(* IEC 61131-3 sources: daoli-st-library/DL_Process (part 70) *)

(* ---- FB_DL_RecipeManager.st ---- *)
(*==============================================================================
 * 组件名称 (Component)  : FB_DL_RecipeManager
 * 所属子库 (Sublibrary) : DL_Process
 * 当前版本 (Version)    : 1.0.1
 * 兼容性 (Platform)   : CODESYS 3.5 / TwinCAT 3 / 汇川 InoProShop / Machine Expert
 *                         仅依赖 Standard.library（R_TRIG），零厂商方言
 * 分类     (Category)   : 工艺段功能块（Function Block · 通用配方管理器）
 * 功能简述 (Function)   : 以「参数清单 + 值集 + 校验和」承载多品种配方：选择、
 *                         校验、应用（写入运行参数）、写回（采集当前参数为
 *                         新配方）、切换防呆（仅机台稳态允许）、变更审计（次
 *                         数 + 注入时间戳）。零文件 I/O、零全局耦合——配方库
 *                         与运行参数均为引脚注入的数组，持久化由调用方自行完
 *                         成；校验和为自包含 32 位滚动异或累加，本块不伪造校
 *                         验和（写回时清零，由调用方重新生成）。
 * 首扫说明 (Init note)  : 纯事件型组件，免首扫（R23/公约 0.1），无 bInit；
 *                         所有状态由指令沿驱动。
 * 公约遵循 (Convention) : 0.2/R21 bError 为显式排除信息级码的派生式；0.4 双语
 *                         同行注释；0.5/R7 实例主体最前部无条件刷新；0.7/R15
 *                         故障锁存仅复位路径清码、信息级瞬时型；0.8 码位段
 *                         16#0005_xxxx（经 DL_Process VERSION.md 复核，本块
 *                         0140~0143 / 0240~0246 无冲突）；0.14 数组存取先判
 *                         域再索引、除法前判零（进度类运算无除法）；0.16 无
 *                         魔法数；0.17 终结符成对 ✓；0.18 ST_DL_RecipeEntry
 *                         与 E_DL_RecipeState 随本块同文件发布；0.19 码位同
 *                         行【级别】注释；0.20 验收向量入头注释；R25 bDone
 *                         单拍生命周期三律。
 * 红线自检 (Redline)    : R1 零全局变量表/外部变量引用 ✓｜R2 零物理 IO 地址 ✓
 *                         R3 纯 IEC 61131-3 ✓｜R4 越界/非有限值/校验和防御 ✓
 *                         R5 全变量中英双语同行注释 ✓｜R6 ENUM+CASE+ELSE ✓
 *                         R7 五实例（R_TRIG×4）主体最前部无条件刷新 ✓
 *                         R8 全常量化 ✓｜R25 单拍标志生命周期三律 ✓
 * 设计要点 (Key notes)  : ① 校验链（eValidating）：配方号域内 → 配方启用 →
 *                           参数个数一致 → 逐参数非有限值 → 逐参数上下限 →
 *                           校验和比对，任一失败锁存对应故障级码；
 *                         ② 应用（eApplying）单拍全量写入 afParamActual，防
 *                           半套参数生效；复核（eVerifying）回读重算校验和比
 *                           对，失败判写入异常 0245；
 *                         ③ 写回（Save）：运行参数拷入配方、个数同步、校验和
 *                           清零（本块不伪造校验和，调用方持久化前须重算）；
 *                         ④ 切换防呆：bMachineStopped=FALSE 时加载拒绝（信
 *                           息码 0141，不置故障，属正常联锁）；Load/Save 同
 *                           拍双丢弃（信息码 0142，"不猜"原则）；
 *                         ⑤ bParamOutOfRange 为瞬时型每拍重算（对当前选中配
 *                           方值集逐参数复核上下限），nOutOfRangeIndex 指向
 *                           首个越界参数；
 *                         ⑥ 数组维度字面量 16（等同 DL_RECIPE_MAX_PARAM）/32
 *                           （等同 DL_RECIPE_MAX_COUNT）与常量同步维护（跨
 *                           平台数组维度须编译期字面量，运行期域检查用常量）。
 * 偏离留档 (Deviation)  : 依 R11 头注释留档，共 1 条：
 *                         ① 校验和算法二选一裁定：规格允许复用 DL_Base 既有
 *                           CRC 函数或自包含算法；本块选自包含 32 位滚动异或
 *                           累加（uSum := (uSum XOR SHL(uSum,5)) +
 *                           REAL_TO_UDINT(v×1000.0 + 1.0E9)，正偏置保证折叠
 *                           项非负、避免负值参数取整的平台回绕歧义；取整语义
 *                           依平台四舍五入）。理由：保持本文件零跨子库依赖，
 *                           可单独导入；影响：与上层持久化校验格式必须一致
 *                           （调用方生成校验和时用同一含偏置算法），头注释已
 *                           声明。
 * 开源溯源 (Origin)     : 来源标签 codesys-forge / recipe-management
 *                         （RAW_NOTES_R8 S-6，T1-4 CODESYS Forge 首次开组：
 *                         公开配方管理示例——配方名/启用/参数值集/校验和的组
 *                         织分类与「校验→应用→复核」相语义，公开开源示例，
 *                         仅借鉴分类与参数域；结构体字段、状态机、码位、引脚
 *                         契约 100% 本库独立设计，clean-room 未复制源码。
 *                         许可证说明：借鉴对象为公开社区示例，本文件为本库原
 *                         创实现，随本库许可证发布）。
 * 验收向量 (Acceptance) :
 *   V1 正常 Load（3 参数，域内）→ bLoaded/eDone、uActiveChecksum 正确、
 *      uChangeCount +1、tLastChange 等于注入 tNow；
 *   V2 参数越界 → 故障 0243 + nOutOfRangeIndex 指向首个越界项；
 *   V3 校验和不匹配 → 0244（配方损坏）；
 *   V4 bMachineStopped=FALSE 加载 → 拒绝 + 信息码 0141（不置故障）；
 *   V5 Save 后 uChangeCount +1、配方值集与个数同步、uChecksum 清零；
 *   V6 Load+Save 同拍 → 双丢弃 + 信息码 0142；
 *   V7 配方参数含非有限值 → 0242；
 *   V8 配方号越界/未启用 → 0240。
 * 修订历史 (Revision)   :
 *   2026-11-15  v1.0.0  首版入库（Round 08 · DL_Process 配方管理件）
 *   2026-11-15  v1.0.1  R8 总监终审修复：终端态分支内的孤立空语句 `;`（非 IEC 61131-3 文法，statement_list 允许零条语句但不容纳孤立分号）改为纯注释占位分支，行为等价、跨平台可移植性合规。
 *============================================================================*)

(*-----------------------------------------------------------------------------
 * 结构体: ST_DL_RecipeEntry（归属 FB_DL_RecipeManager，与其同文件发布）
 *         值集维度字面量 16 等同 DL_RECIPE_MAX_PARAM，须与常量同步维护。
 *----------------------------------------------------------------------------*)
TYPE ST_DL_RecipeEntry :
STRUCT
    sName        : STRING[32];                    // 配方名（Recipe name）/ Recipe name
    bEnabled     : BOOL;                          // 配方启用（Enabled），FALSE 时选中即判故障 / Recipe enabled flag
    nParamCount  : UINT;                          // 有效参数个数（Active param count）[-]，域 0..16 / Active parameter count
    afValue      : ARRAY[0..15] OF REAL;          // 参数值集（Parameter values），维度 16 等同 DL_RECIPE_MAX_PARAM / Parameter values, dim 16
    uChecksum    : UDINT;                         // 校验和（Checksum），0=未启用校验；由调用方生成、本块只比对 / Checksum, 0 = verification off, caller generates
END_STRUCT
END_TYPE

(*-----------------------------------------------------------------------------
 * 枚举: E_DL_RecipeState（归属 FB_DL_RecipeManager，与其同文件发布）
 *----------------------------------------------------------------------------*)
TYPE E_DL_RecipeState :
(
    eIdle       := 0,   // 空闲：等操作沿 / Idle, awaiting operation edge
    eValidating := 10,  // 校验中：选择域/启用/个数/数值域/校验和逐项过链 / Validating selection, enable, count, ranges and checksum
    eApplying   := 20,  // 应用中：加载全量写入运行参数 / 写回采集参数入配方 / Applying, load writes parameters or save collects them
    eVerifying  := 30,  // 复核中：回读运行参数重算校验和比对 / Verifying, read-back checksum comparison
    eDone       := 40,  // 完成：结果保持，等下一操作沿 / Done, results held awaiting next operation
    eFault      := 99   // 故障锁存：仅复位沿退出 / Fault latched, only reset edge exits
) UINT;
END_TYPE

FUNCTION_BLOCK FB_DL_RecipeManager
VAR_INPUT
    bEnable             : BOOL;             // 使能（Enable），FALSE=中止操作并保持当前运行参数不变 / Enable, FALSE aborts and keeps live parameters
    bLoad               : BOOL;             // 加载所选配方到运行参数（Load），上升沿受理 / Load edge applies selected recipe
    bSave               : BOOL;             // 把当前运行参数写回所选配方（Save/Teach），上升沿受理 / Save edge teaches live parameters into recipe
    bValidate           : BOOL;             // 仅校验不应用（Validate），上升沿受理，结果出 bValid / Validate edge, result in bValid
    bMachineStopped     : BOOL := TRUE;     // 机台稳态确认（Machine stopped），FALSE 时拒绝加载（切换防呆）/ Machine stopped interlock, FALSE rejects load
    bReset              : BOOL;             // 复位故障（Fault reset），上升沿受理 / Rising edge resets fault
    nSelectRecipe       : UINT;             // 选中配方号（Selected recipe index）[-]，域 0..DL_RECIPE_MAX_COUNT-1 / Selected recipe index
    nParamCount         : UINT := 1;        // 本机参数个数（Param count）[-]，域 1..DL_RECIPE_MAX_PARAM，越界钳位 / Machine parameter count, clamped
    afParamMin          : ARRAY[0..15] OF REAL; // 参数下限（Param lower limits），逐项与配方值比较；min ≥ max 视为该参数未启用校验 / Param lower limits, min ≥ max disables that check
    afParamMax          : ARRAY[0..15] OF REAL; // 参数上限（Param upper limits），与下限配对使用 / Param upper limits paired with lower
    tNow                : TIME := T#0S;     // 时间戳注入（Timestamp injection）[ms]，禁读 CPU 钟，用于审计记录 / Injected timestamp for audit, CPU clock never read
END_VAR
VAR_OUTPUT
    bLoaded             : BOOL;             // 加载完成（Loaded），完成态且操作为 Load 时为 TRUE / TRUE while done with load operation
    bSaved              : BOOL;             // 写回完成（Saved），完成态且操作为 Save 时为 TRUE / TRUE while done with save operation
    bValid              : BOOL;             // 校验通过（Valid），校验型操作结果，保持到下次操作 / Validation verdict held until next operation
    bParamOutOfRange    : BOOL;             // 存在越界参数（Out of range），瞬时型每拍重算 / Transient out-of-range flag, recomputed each scan
    nOutOfRangeIndex    : UINT;             // 首个越界参数索引（First bad index）[-]，越界标志有效时成立 / First out-of-range parameter index
    nActiveRecipe       : UINT;             // 当前生效配方号（Active recipe）[-] / Currently applied recipe index
    uActiveChecksum     : UDINT;            // 当前运行参数校验和（Active checksum），每拍重算供上层比对 / Live parameter checksum recomputed each scan
    uChangeCount        : UDINT;            // 配方变更次数（Change counter），每次成功 Load/Save +1 / Successful load/save counter
    tLastChange         : TIME := T#0S;     // 末次变更时间戳（Last change time），取注入 tNow / Last change timestamp from injected tNow
    bBusy               : BOOL;             // 执行中（Busy），校验/应用/复核态为 TRUE / TRUE while validating/applying/verifying
    bDone               : BOOL;             // 操作完成单拍脉冲（Done pulse），单拍生命周期三律 / One-scan operation done pulse
    bError              : BOOL;             // 故障锁存（Error），仅故障级码置位 / Latched error, fault codes only
    uErrorId            : UDINT;            // 故障码（Error code），16#0005_xxxx 段，0=无故障 / Error code, fault-level priority
END_VAR
VAR_IN_OUT
    astRecipe           : ARRAY[0..31] OF ST_DL_RecipeEntry; // 配方库（Recipe library），维度 32 等同 DL_RECIPE_MAX_COUNT，调用方持有与持久化 / Recipe library owned and persisted by caller
    afParamActual       : ARRAY[0..15] OF REAL; // 当前运行参数（Live parameters），维度 16，Save 被读 / Load 被写 / Live parameters, read on save, written on load
END_VAR
VAR
    _eState             : E_DL_RecipeState := E_DL_RecipeState.eIdle; // 内部状态机（Internal state）/ Internal state
    _nOp                : USINT;            // 当前操作类型（Operation type）[-]，1=Load 2=Save 3=Validate，0=无 / Operation type register
    _bFaultLatch        : BOOL;             // 故障锁存标志（Fault latch flag），仅复位路径清除 / Fault latch, cleared only via reset path
    _uErrorIdInt        : UDINT;            // 内部故障级码寄存（Internal fault-level register）/ Internal fault-level register
    _uInfoCode          : UDINT;            // 本拍信息级码（Info code this cycle），瞬时型每拍重算 / Transient info code
    _nParamEff          : UINT;             // 生效参数个数（Effective param count），钳位后值 / Clamped effective parameter count
    _nSelEff            : UINT;             // 生效配方号（Effective recipe index），域校验后值 / Validated recipe index
    _fV                 : REAL;             // 循环内当前参数值（Loop value scratch）/ Loop parameter value scratch
    _bFinite            : BOOL;             // 非有限值检测结果（Finite check verdict）/ Finite-value check verdict
    _uSum               : UDINT;            // 校验和累加器（Checksum accumulator）/ Checksum accumulator
    _uTargetCk          : UDINT;            // 目标配方校验和（Target recipe checksum）/ Target recipe checksum
    _nIdx               : UINT;             // 循环索引（Loop index）[-] / Loop index
    _bBadIdxFound       : BOOL;             // 越界首索引已记录（First bad index found）/ First bad index recorded flag
    _bValOk             : BOOL;             // 校验链通过（Validation chain passed）/ Validation chain verdict
    _fbTrigLoad         : R_TRIG;           // 加载沿（Load edge detector）/ Load edge detector
    _fbTrigSave         : R_TRIG;           // 写回沿（Save edge detector）/ Save edge detector
    _fbTrigValidate     : R_TRIG;           // 校验沿（Validate edge detector）/ Validate edge detector
    _fbTrigReset        : R_TRIG;           // 复位沿（Reset edge detector）/ Reset edge detector
END_VAR
VAR CONSTANT
    DL_RECIPE_MAX_PARAM : UINT := 16;       // 单配方参数上限（Max params per recipe）[-]，与数组维度字面量 16 同步 / Max params, sync with literal dim 16
    DL_RECIPE_MAX_COUNT : UINT := 32;       // 配方库容量上限（Max recipe count）[-]，与数组维度字面量 32 同步 / Max recipes, sync with literal dim 32
    DL_RECIPE_REAL_MAX  : REAL := 3.4E38;   // 单精度有限值判据幅值（Finite magnitude bound），超出或非数均拒绝 / Finite magnitude bound for REAL inputs
    DL_RECIPE_EPS       : REAL := 1.0E-6;   // 浮点通用容差（General float epsilon）/ General float epsilon
    DL_RECIPE_VERIFY_EPS: REAL := 1.0E-3;   // 复核逐参数容差（Verify per-param epsilon），千分之一工程单位 / Verify tolerance per parameter
    DL_RECIPE_SCALE     : REAL := 1000.0;   // 校验和定标系数（Checksum scale）[-]，值×此系数取整入校验和 / Checksum scale factor for fixed-point fold
    DL_RECIPE_BIAS      : REAL := 1.0E9;    // 校验和正偏置（Checksum positive bias），保证折叠项非负、跨平台回绕确定 / Positive bias keeps fold term non-negative, portable
    DL_RECIPE_CHK_ROL   : DINT := 5;        // 校验和滚动移位量（Checksum shift amount）[-] / Checksum rolling shift amount
    DL_RECIPE_OP_LOAD   : USINT := 1;       // 操作码：加载（Op code: load）/ Op code load
    DL_RECIPE_OP_SAVE   : USINT := 2;       // 操作码：写回（Op code: save）/ Op code save
    DL_RECIPE_OP_VALID  : USINT := 3;       // 操作码：仅校验（Op code: validate only）/ Op code validate-only
    DL_RECIPE_ERR_SEL   : UDINT := 16#0005_0240; // 0005_0240 配方号越界/未启用【故障级】/ Bad recipe index or disabled, fault level
    DL_RECIPE_ERR_CNT   : UDINT := 16#0005_0241; // 0005_0241 参数个数与配方定义不一致【故障级】/ Param count mismatch, fault level
    DL_RECIPE_ERR_NAN   : UDINT := 16#0005_0242; // 0005_0242 配方参数含非有限值【故障级】/ Non-finite recipe parameter, fault level
    DL_RECIPE_ERR_RANGE : UDINT := 16#0005_0243; // 0005_0243 参数越界【故障级】/ Parameter out of range, fault level
    DL_RECIPE_ERR_CKSUM : UDINT := 16#0005_0244; // 0005_0244 校验和不匹配（配方损坏）【故障级】/ Checksum mismatch, recipe corrupted, fault level
    DL_RECIPE_ERR_VERIFY: UDINT := 16#0005_0245; // 0005_0245 应用后复核失败【故障级】/ Post-apply verify failed, fault level
    DL_RECIPE_ERR_STATE : UDINT := 16#0005_0246; // 0005_0246 非法状态兜底【故障级】/ Illegal state fallback, fault level
    DL_RECIPE_INFO_NOCK : UDINT := 16#0005_0140; // 0005_0140 配方未启用校验和（uChecksum=0）【信息级】/ Checksum disabled (zero), info level
    DL_RECIPE_INFO_LOCK : UDINT := 16#0005_0141; // 0005_0141 机台非稳态，加载被拒【信息级】/ Load rejected, machine not stopped, info level
    DL_RECIPE_INFO_CONF : UDINT := 16#0005_0142; // 0005_0142 Load/Save 同拍冲突，双丢弃【信息级】/ Load/save edge conflict, both dropped, info level
    DL_RECIPE_INFO_CLAMP: UDINT := 16#0005_0143; // 0005_0143 参数个数越界钳位【信息级】/ Param count clamped, info level
END_VAR

// ============================================================================
// 段 1｜实例无条件周期刷新（R7/0.5：严禁置于 IF/CASE 分支内）
//      Unconditional per-cycle refresh of all instances (R7/0.5)
// ============================================================================
_fbTrigLoad(CLK := bLoad);              // 加载沿（Load edge）
_fbTrigSave(CLK := bSave);              // 写回沿（Save edge）
_fbTrigValidate(CLK := bValidate);      // 校验沿（Validate edge）
_fbTrigReset(CLK := bReset);            // 复位沿（Reset edge）

// ============================================================================
// 段 2｜信息级预清零 + 单拍标志预清零 + 参数防御（R25/R15）
//      Info preset + one-shot preset + parameter defense (R25/R15)
// ============================================================================
_uInfoCode := 0;                        // 信息级瞬时型每拍重算（Transient info recomputed each scan）
bDone := FALSE;                         // 完成单拍先清零（R25：置位-消费-复位同周期闭环）/ Done pulse preset FALSE (R25 lifecycle)

// 参数个数钳位（Param count clamp，域 1..16）
IF nParamCount < UINT#1 THEN
    _nParamEff := UINT#1;               // 下限钳位（Lower clamp）
    _uInfoCode := DL_RECIPE_INFO_CLAMP; // 0005_0143 参数个数越界钳位【信息级】/ Count clamped, info level
ELSIF nParamCount > DL_RECIPE_MAX_PARAM THEN
    _nParamEff := DL_RECIPE_MAX_PARAM;  // 上限钳位（Upper clamp）
    _uInfoCode := DL_RECIPE_INFO_CLAMP; // 0005_0143 参数个数越界钳位【信息级】/ Count clamped, info level
ELSE
    _nParamEff := nParamCount;          // 引脚原值（Pin value as-is）
END_IF

// 复位路径：仅此路径可清故障锁存（R15）
IF _fbTrigReset.Q THEN
    _bFaultLatch := FALSE;              // 故障锁存解除（Fault latch released）
    _uErrorIdInt := 16#0000_0000;       // 故障码清零（Fault code cleared）
    IF _eState = E_DL_RecipeState.eFault THEN
        _eState := E_DL_RecipeState.eIdle; // 故障态回空闲（Fault state back to idle）
    END_IF
END_IF

// ============================================================================
// 段 3｜每拍瞬态复核：运行参数校验和 + 越界扫描（对当前选中配方）
//      Per-scan transient: live checksum + out-of-range scan on selected recipe
// ============================================================================
uActiveChecksum := 16#0000_0000;        // 校验和累加器清零（Checksum accumulator reset）
FOR _nIdx := UINT#0 TO _nParamEff - UINT#1 DO
    _fV := afParamActual[_nIdx];        // 索引域已由 _nParamEff 钳位保证（Index bounded by clamped count）
    uActiveChecksum := (uActiveChecksum XOR SHL(uActiveChecksum, DL_RECIPE_CHK_ROL))
                  + REAL_TO_UDINT(_fV * DL_RECIPE_SCALE + DL_RECIPE_BIAS);   // 滚动异或累加 + 正偏置保证非负折叠（偏离留档①算法）/ Rolling XOR fold with positive bias (deviation 1)
END_FOR

bParamOutOfRange := FALSE;              // 越界标志瞬态预清零（Transient flag preset）
nOutOfRangeIndex := UINT#0;             // 首个越界索引预清零（First bad index preset）
IF nSelectRecipe < DL_RECIPE_MAX_COUNT THEN
    IF (astRecipe[nSelectRecipe].nParamCount >= UINT#1)
      AND (astRecipe[nSelectRecipe].nParamCount <= DL_RECIPE_MAX_PARAM) THEN
        FOR _nIdx := UINT#0 TO astRecipe[nSelectRecipe].nParamCount - UINT#1 DO
            _fV := astRecipe[nSelectRecipe].afValue[_nIdx];      // 配方值（Recipe value）
            IF (afParamMin[_nIdx] < afParamMax[_nIdx])
              AND ((_fV < afParamMin[_nIdx]) OR (_fV > afParamMax[_nIdx]))
              AND (NOT bParamOutOfRange) THEN
                bParamOutOfRange := TRUE;            // 越界成立（Out of range found）
                nOutOfRangeIndex := _nIdx;           // 首个越界索引（First bad index）
            END_IF
        END_FOR
    END_IF
END_IF

// ============================================================================
// 段 4｜操作受理（仅在空闲/完成态受理指令沿；同拍冲突双丢弃）
//      Operation acceptance at idle/done; same-cycle conflict drops both
// ============================================================================
IF bEnable AND (( _eState = E_DL_RecipeState.eIdle)
             OR (_eState = E_DL_RecipeState.eDone)) THEN
    IF _fbTrigLoad.Q AND _fbTrigSave.Q THEN
        _uInfoCode := DL_RECIPE_INFO_CONF;  // 0005_0142 Load/Save 同拍冲突双丢弃【信息级】/ Edge conflict, both dropped
    ELSIF _fbTrigLoad.Q THEN
        IF bMachineStopped THEN
            _nOp := DL_RECIPE_OP_LOAD;      // 登记加载操作（Register load operation）
            _eState := E_DL_RecipeState.eValidating;
        ELSE
            _uInfoCode := DL_RECIPE_INFO_LOCK; // 0005_0141 机台非稳态加载被拒【信息级】/ Load rejected, machine running
        END_IF
    ELSIF _fbTrigSave.Q THEN
        _nOp := DL_RECIPE_OP_SAVE;          // 登记写回操作（Register save operation）
        _eState := E_DL_RecipeState.eValidating;
    ELSIF _fbTrigValidate.Q THEN
        _nOp := DL_RECIPE_OP_VALID;         // 登记校验操作（Register validate operation）
        _eState := E_DL_RecipeState.eValidating;
    END_IF
END_IF

// ============================================================================
// 段 5｜核心状态机（ENUM + CASE，含 ELSE 非法状态兜底）
//      Core state machine (ENUM + CASE with ELSE fallback)
// ============================================================================
CASE _eState OF

    E_DL_RecipeState.eIdle: // 空闲：等操作沿（受理逻辑在段 4）
        // 无动作（No action）

    E_DL_RecipeState.eValidating: // 校验链：域 → 启用 → 个数 → 非有限值 → 上下限 → 校验和
        _bValOk := TRUE;                    // 校验链初始通过（Chain starts valid）
        // ① 配方号域内（Index in domain）
        IF nSelectRecipe >= DL_RECIPE_MAX_COUNT THEN
            _bValOk := FALSE;
            _bFaultLatch := TRUE;
            _uErrorIdInt := DL_RECIPE_ERR_SEL;   // 0005_0240 配方号越界【故障级】/ Bad recipe index, fault level
        ELSE
            _nSelEff := nSelectRecipe;           // 生效配方号登记（Register effective index）
            // ② 配方启用（Recipe enabled）
            IF NOT astRecipe[_nSelEff].bEnabled THEN
                _bValOk := FALSE;
                _bFaultLatch := TRUE;
                _uErrorIdInt := DL_RECIPE_ERR_SEL; // 0005_0240 配方未启用【故障级】/ Recipe disabled, fault level
            END_IF
        END_IF

        IF _bValOk THEN
            // ③ 参数个数一致（Load/Validate 要求；Save 允许覆盖定义）
            IF (_nOp <> DL_RECIPE_OP_SAVE)
              AND (astRecipe[_nSelEff].nParamCount <> _nParamEff) THEN
                _bValOk := FALSE;
                _bFaultLatch := TRUE;
                _uErrorIdInt := DL_RECIPE_ERR_CNT;   // 0005_0241 个数与配方定义不一致【故障级】/ Count mismatch, fault level
            END_IF
        END_IF

        IF _bValOk AND (_nOp <> DL_RECIPE_OP_SAVE) THEN
            _uTargetCk := 16#0000_0000;          // 目标校验和累加器（Target checksum accumulator）
            FOR _nIdx := UINT#0 TO _nParamEff - UINT#1 DO
                _fV := astRecipe[_nSelEff].afValue[_nIdx];    // 配方值（Recipe value）
                _bFinite := (_fV >= (-DL_RECIPE_REAL_MAX)) AND (_fV <= DL_RECIPE_REAL_MAX); // 非有限值自比等价式（Finite check）
                IF NOT _bFinite THEN
                    _bValOk := FALSE;
                    _bFaultLatch := TRUE;
                    _uErrorIdInt := DL_RECIPE_ERR_NAN;        // 0005_0242 参数含非有限值【故障级】/ Non-finite parameter, fault level
                ELSIF (afParamMin[_nIdx] < afParamMax[_nIdx])
                  AND ((_fV < afParamMin[_nIdx]) OR (_fV > afParamMax[_nIdx])) THEN
                    _bValOk := FALSE;
                    _bFaultLatch := TRUE;
                    _uErrorIdInt := DL_RECIPE_ERR_RANGE;      // 0005_0243 参数越界【故障级】/ Parameter out of range, fault level
                    nOutOfRangeIndex := _nIdx;                // 首个越界索引（First bad index）
                END_IF
                _uTargetCk := (_uTargetCk XOR SHL(_uTargetCk, DL_RECIPE_CHK_ROL))
                         + REAL_TO_UDINT(_fV * DL_RECIPE_SCALE + DL_RECIPE_BIAS);   // 同算法重算目标校验和（Target checksum recomputed, same algorithm）
            END_FOR
            // ⑤ 校验和比对（=0 视为未启用校验）
            IF _bValOk THEN
                IF astRecipe[_nSelEff].uChecksum = 16#0000_0000 THEN
                    _uInfoCode := DL_RECIPE_INFO_NOCK;    // 0005_0140 未启用校验和【信息级】/ Checksum disabled, info level
                ELSIF astRecipe[_nSelEff].uChecksum <> _uTargetCk THEN
                    _bValOk := FALSE;
                    _bFaultLatch := TRUE;
                    _uErrorIdInt := DL_RECIPE_ERR_CKSUM;  // 0005_0244 校验和不匹配（配方损坏）【故障级】/ Checksum mismatch, fault level
                END_IF
            END_IF
        END_IF

        // 校验链出口分派（Chain exit dispatch）
        IF _bValOk THEN
            IF _nOp = DL_RECIPE_OP_LOAD THEN
                _eState := E_DL_RecipeState.eApplying;    // 进入应用（Proceed to apply）
            ELSIF _nOp = DL_RECIPE_OP_SAVE THEN
                _eState := E_DL_RecipeState.eApplying;    // 写回也走应用相（Save proceeds to apply phase）
            ELSE
                bValid := TRUE;                           // 仅校验：结果通过（Validate-only passed）
                bDone := TRUE;                            // 完成单拍（R25 本拍闭环）/ Done pulse (R25)
                _eState := E_DL_RecipeState.eDone;
            END_IF
        ELSE
            _eState := E_DL_RecipeState.eFault;           // 校验失败进故障锁存（Validation failed, latch fault）
        END_IF

    E_DL_RecipeState.eApplying: // 应用：Load 单拍全量写入 / Save 单拍全量采集
        IF _nOp = DL_RECIPE_OP_LOAD THEN
            FOR _nIdx := UINT#0 TO _nParamEff - UINT#1 DO
                _fV := astRecipe[_nSelEff].afValue[_nIdx];    // 源：配方值（Source: recipe value）
                _bFinite := (_fV >= (-DL_RECIPE_REAL_MAX)) AND (_fV <= DL_RECIPE_REAL_MAX);
                IF _bFinite THEN
                    afParamActual[_nIdx] := _fV;              // 单拍全量写入（Single-scan bulk write, no half-set applied）
                END_IF
            END_FOR
            _eState := E_DL_RecipeState.eVerifying;           // 进入复核（Proceed to verify）
        ELSE
            FOR _nIdx := UINT#0 TO _nParamEff - UINT#1 DO
                astRecipe[_nSelEff].afValue[_nIdx] := afParamActual[_nIdx]; // 单拍全量采集（Single-scan bulk collect）
            END_FOR
            astRecipe[_nSelEff].nParamCount := _nParamEff;    // 个数同步（Count synchronized）
            astRecipe[_nSelEff].uChecksum := 16#0000_0000;    // 校验和清零：本块不伪造，调用方须重算（Checksum zeroed, caller regenerates）
            uChangeCount := uChangeCount + UINT#1;            // 审计计数（Audit counter）
            tLastChange := tNow;                              // 审计时间戳取注入值（Audit timestamp from injected pin）
            nActiveRecipe := _nSelEff;                        // 生效配方号登记（Active recipe registered）
            bSaved := TRUE;                                   // 写回完成保持（Saved held）
            bDone := TRUE;                                    // 完成单拍（R25 本拍闭环）/ Done pulse (R25)
            _eState := E_DL_RecipeState.eDone;
        END_IF

    E_DL_RecipeState.eVerifying: // 复核：回读运行参数与目标比对（防写入异常）
        IF astRecipe[_nSelEff].uChecksum <> 16#0000_0000 THEN
            IF uActiveChecksum <> astRecipe[_nSelEff].uChecksum THEN
                _bFaultLatch := TRUE;
                _uErrorIdInt := DL_RECIPE_ERR_VERIFY;         // 0005_0245 复核失败（写入异常）【故障级】/ Verify failed, fault level
                _eState := E_DL_RecipeState.eFault;
            ELSE
                nActiveRecipe := _nSelEff;                    // 生效配方号登记（Active recipe registered）
                uChangeCount := uChangeCount + UINT#1;        // 审计计数（Audit counter）
                tLastChange := tNow;                          // 审计时间戳（Audit timestamp）
                bLoaded := TRUE;                              // 加载完成保持（Loaded held）
                bDone := TRUE;                                // 完成单拍（R25 本拍闭环）/ Done pulse (R25)
                _eState := E_DL_RecipeState.eDone;
            END_IF
        ELSE
            // 目标未启用校验和：逐参数容差比对兜底（Checksum off: element-wise tolerance fallback）
            FOR _nIdx := UINT#0 TO _nParamEff - UINT#1 DO
                IF ABS(afParamActual[_nIdx] - astRecipe[_nSelEff].afValue[_nIdx]) > DL_RECIPE_VERIFY_EPS THEN
                    _bFaultLatch := TRUE;
                    _uErrorIdInt := DL_RECIPE_ERR_VERIFY;     // 0005_0245 复核失败【故障级】/ Verify failed, fault level
                    _eState := E_DL_RecipeState.eFault;
                END_IF
            END_FOR
            IF NOT _bFaultLatch THEN
                nActiveRecipe := _nSelEff;
                uChangeCount := uChangeCount + UINT#1;
                tLastChange := tNow;
                bLoaded := TRUE;                              // 加载完成保持（Loaded held）
                bDone := TRUE;                                // 完成单拍（R25）/ Done pulse (R25)
                _eState := E_DL_RecipeState.eDone;
            END_IF
        END_IF

    E_DL_RecipeState.eDone: // 完成：结果保持，下一操作沿回空闲（受理逻辑在段 4，下一拍起效）
        IF _fbTrigLoad.Q OR _fbTrigSave.Q OR _fbTrigValidate.Q THEN
            _eState := E_DL_RecipeState.eIdle;                // 让位新操作（Yield to new operation）
            bLoaded := FALSE;                                 // 结果锁存随让位清零（Result holds released）
            bSaved := FALSE;
            bValid := FALSE;
        END_IF

    E_DL_RecipeState.eFault: // 故障锁存：等复位（复位路径在段 2）
        // 等复位（Awaiting reset）

    ELSE // 非法状态兜底（本块专用码位）
        _bFaultLatch := TRUE;
        _uErrorIdInt := DL_RECIPE_ERR_STATE;                  // 0005_0246 非法状态兜底【故障级】/ Illegal state fallback, fault level
        _eState := E_DL_RecipeState.eFault;
END_CASE

// ============================================================================
// 段 6｜使能撤销与出口派生（R21）
//      Enable teardown and outlet derivation (R21)
// ============================================================================
IF NOT bEnable THEN
    // 撤销进行中操作，运行参数保持不变（Abort in-flight ops, live parameters untouched）
    IF (_eState = E_DL_RecipeState.eValidating)
     OR (_eState = E_DL_RecipeState.eApplying)
     OR (_eState = E_DL_RecipeState.eVerifying) THEN
        _eState := E_DL_RecipeState.eIdle;   // 中途回空闲（Back to idle mid-flight）
    END_IF
END_IF

bBusy := (_eState = E_DL_RecipeState.eValidating)
      OR (_eState = E_DL_RecipeState.eApplying)
      OR (_eState = E_DL_RecipeState.eVerifying);            // 执行中派生（Busy derived）

bError := _bFaultLatch;                      // 故障级派生式（Fault-level derived form）
IF _bFaultLatch THEN
    uErrorId := _uErrorIdInt;                // 故障级码优先透出（Fault-level priority）
ELSE
    uErrorId := _uInfoCode;                  // 无故障时透出本拍信息级码（Transient info code）
END_IF
END_FUNCTION_BLOCK

(* ---- FB_DL_RejectBlowCtrl.st ---- *)
(*
    FB_DL_RejectBlowCtrl —— 输送线剔除气吹执行时序（NG 预告 → 距离/速度延时 → 定宽气吹 → 对账）
    ------------------------------------------------------------------
    组件名称  : FB_DL_RejectBlowCtrl
    分类      : DL_Process / Rejection
    前缀      : FB_DL_
    版本      : 1.0.0
    溯源      : 自研线 s9-conv（R7 先例同口径）：剔除气吹执行时序属输送线
                工程惯例的 clean-room 自有实现；判定域（视觉 / 称重）与
                诊断域（堵塞）归邻件，本件零借用；实现 / 引脚名 / 码位 /
                对账口径 100% 自有；无闭源参考。
    平台      : 纯 IEC 61131-3（ENUM + CASE + TON / R_TRIG + 标准换算），
                CODESYS 3.5 / TwinCAT 3 / InoProShop / Machine Expert 通用
    作者      : 道莅代码库 · PLC编程专家（R72 构建轮 · 批 4 · 序号 11）
    ------------------------------------------------------------------
    功能说明  : 灌装 / 包装线吹除 NG 瓶：eIdle →（bNgFlag 上升沿布防）
                eArm（延时窗 = fDistNgToGate / fBeltVel 秒换算毫秒，组态
                容差即引脚侧自行加权，本件按纯行程 / 速度口径）→ eBlow
                （定宽气吹脉冲 tBlowPulse）→ eConfirm（确认窗 tConfirmWin
                满拍**复验一次** NG 离线状态，R41/R42 同拍竞态口径：窗满拍
                反馈迟到临界收敛以窗满拍采样为准）→ eIdle。
                对账口径（漏剔 / 误剔 / 剔除三值互斥，窗满拍一次性判归）：
                ① 漏剔 uMissCount：窗满拍 bNgFlag 仍在位（气吹未吹走 NG）；
                ② 误剔 uFalseCount：布防后气吹执行拍 bNgFlag 已离线（无 NG
                   确认却执行气吹——预告为伪沿，好品被吹）；
                ③ 剔除 uRejectCount：气吹拍 NG 在位且窗满拍已离线（正常剔除）。
                漏剔 / 误剔计数直接进 OEE 质量因子。
                安全口径：
                ① fBeltVel 非有限 / <= 0 → **拒收布防 + NG 漏剔计数**（不发
                   气吹，防静默放行——速度不明即不剔除，宁可人工清台），
                   信息级；执行中途速度失效同样撤销布防 + 漏剔计数；
                ② 除法先判后除：fDistNgToGate / fBeltVel 仅在速度过闸后执行；
                   毫秒换算 LREAL→DINT 前做实数上界钳制（DL_RBC_TMAX，
                   防溢出方向翻转，R151）；
                ③ 失能 → bBlowCmd 清零 + 布防撤销（停机相输出清零，R57）；
                   计数保留（OEE 台账语义）；
                ④ 组态闸：tBlowPulse / tConfirmWin 非正 或 fDistNgToGate
                   非有限 / 非正 → 故障锁存（锁存期 NG 沿一律按漏剔计数，
                   宁多计不漏计）。
    错误码    : 16#0005_0630 速度不明拒剔（fBeltVel 非有限 / 非正，布防撤销
                            + 漏剔计数），条件期重算 —— 信息级，不置 bError
                16#0005_0631 组态非法（tBlowPulse / tConfirmWin 非正 /
                            fDistNgToGate 非有限 / 非正），锁存至复位沿
                            —— 故障级
                加码反证句（R90）：0630 由「布防撤销 + 漏剔计数递增」唯一
                观测（正常剔除路径漏剔计数不动）；0631 与 0630 输出可分
                （bError 与锁存回放 vs 条件信息级），成因互斥（组态表 vs
                运行速度），故各立一码。
    码位总账  : 16#0005_0630 用 ｜ 16#0005_0631 用
                （0620~0622 / 3036~3038 已由同段邻件占用，本件不占）
    边界与披露: 一 R_TRIG（rtNg / rtReset）与 TON（tonPhase）每拍**无条件
                   调用**（规则 ⑦）；tonPhase PT 按相选择（布防延时 / 气吹
                   定宽 / 确认窗三态一实例，R367 逐相 PT 口径），IN = 相驻留
                   显式变量；
                二 零全局变量、零 VAR_EXTERNAL、零物理地址；
                三 归属 Ownership：E_DL_RejectPhase 属主为本文件（全库唯一
                   定义，R264），引用件只引用不重声明；
                四 状态机 ENUM + CASE 必带 ELSE 兜底（非法枚举值 → eFault
                   锁存）+ 段 5b 统一故障迁入闸（R274）；
                五 域闸逐项点名（R272）：fBeltVel / fDistNgToGate 双浮点引脚
                   全部纳入非有限与符号闸；
                六 换算链：tArmDelay := DINT_TO_TIME(LREAL_TO_DINT(钳制后的
                   行程毫秒))，钳制上界 2147483000 ms（< 2^31 − 347，
                   LREAL_TO_DINT 域内可表反算，R63）；
                七 分工声明：FB_DL_VisionResultGate（视觉结果放行闸）、
                   FB_DL_WeightCheckReject（称重 NG 判定）、
                   FB_DL_ConveyorJamDetect（堵塞诊断）——三者均属「判定」域，
                   本件只做「预告 → 延时 → 气吹 → 对账」**执行时序**域
                   （R363 邻接共存先例），不判 NG、不诊断堵塞；
                八 复位沿作用域（R311）：清故障锁存 + 清锁存码 + 迁 eIdle +
                   撤布防，**不清** uRejectCount / uMissCount / uFalseCount
                   （OEE 台账语义，只随失能保留、由上位归档后清）；
                九 依赖声明：仅 Standard.library（TON / R_TRIG），零厂商
                   方言；
                十 接口契约：bNgFlag 须为**电平型**预告（预告对象离线前保持
                   在位），脉型预告会在气吹拍被判为误剔（uFalseCount 虚高）
                   ——脉型上游须先展宽再接入；失能相（bEn = FALSE）的 NG 沿
                   不布防不计数（停线工况，宁缺勿滥口径）。
    验收向量  : V1 正常剔除：NG 沿 → 行程延时 → 气吹拍 NG 在位 → 窗满拍
                NG 离线 → uRejectCount + 1；
                V2 漏剔：窗满拍 bNgFlag 仍在位 → uMissCount + 1；
                V3 误剔：气吹拍 bNgFlag 已离线 → uFalseCount + 1；
                V4 fBeltVel = 0 / NaN → NG 沿按漏剔计数、不发气吹、0630；
                V5 tBlowPulse = T#0MS → 0631 锁存；V6 失能 → bBlowCmd 清零
                + 布防撤销；V7 复位沿 → 解锁回 eIdle（计数不清）。
                算法已证（脚本）：未跑 ｜ 编译器已证（三平台）：未跑
    修订记录  : 2026-11-23 v1.0.0 首次入库（R72 构建轮 · 批 4 · 序号 11）
*)
TYPE E_DL_RejectPhase :
(
    eIdle    := 0,                         // 空闲：等 NG 预告沿布防 / idle, waiting for the NG leading edge
    eArm     := 10,                        // 布防延时：行程 / 速度换算延时窗 / armed, the travel delay window
    eBlow    := 20,                        // 定宽气吹：tBlowPulse 定宽脉冲 / blowing, the fixed width pulse
    eConfirm := 30,                        // 确认窗：窗满拍复验 NG 离线 / confirm, the recheck window
    eFault   := 60                         // 故障：锁存待复位 / fault, latched until the reset
);
END_TYPE

FUNCTION_BLOCK FB_DL_RejectBlowCtrl
VAR_INPUT
    bNgFlag       : BOOL := FALSE;         (* 上游 NG 预告（视觉 / 称重判定输出），[标志] / the upstream NG leading flag *)
    fBeltVel      : LREAL := 1000.0;       (* 输送带速度，[mm/s]，非有限或非正拒剔 / the belt velocity in mm per second *)
    fDistNgToGate : LREAL := 500.0;        (* NG 检测位到气吹位间距，[mm]，禁非有限 / 非正 / the distance from the detector to the gate in mm *)
    tBlowPulse    : TIME := T#100MS;       (* 气吹定宽，[ms]，禁非正 / the blow pulse width *)
    tConfirmWin   : TIME := T#200MS;       (* 剔除确认窗，[ms]，禁非正 / the reject confirmation window *)
    bEn           : BOOL := FALSE;         (* 使能，[标志]，FALSE 撤布防清气吹（计数保留）/ the enable *)
    bReset        : BOOL := FALSE;         (* 故障复位，[标志]，上升沿唯一解除 / the fault reset *)
END_VAR
VAR_OUTPUT
    bBlowCmd    : BOOL := FALSE;           (* 气吹指令出口（定宽脉冲），[标志] / the blow command outlet *)
    uRejectCount: UDINT := 0;              (* 剔除成功计数（OEE 台账），[件] / the successful reject count *)
    uMissCount  : UDINT := 0;              (* 漏剔计数（窗满 NG 仍在位 / 速度不明拒剔），[件] / the miss count *)
    uFalseCount : UDINT := 0;              (* 误剔计数（气吹拍 NG 已离线），[件] / the false reject count *)
    eState      : E_DL_RejectPhase := E_DL_RejectPhase.eIdle; // 主状态机当前态 [状态] / the current state
    bError      : BOOL := FALSE;           (* 故障标志，与锁存同源（R191）/ the fault flag from the latch *)
    nErrCode    : UDINT := 16#0000_0000;   (* 错误码，0 = 正常，故障锁存回放（R187）/ the error id *)
END_VAR
VAR
    _bInit      : BOOL := FALSE;           (* 首拍初始化标志（R310）/ the first scan flag *)
    _eState     : E_DL_RejectPhase := E_DL_RejectPhase.eIdle; // 内部状态寄存器 / the internal state register
    _bFault     : BOOL := FALSE;           (* 故障锁存副本，仅复位沿解除 / the fault latch copy *)
    _nCodeLatch : UDINT := 0;              (* 锁存成因码，故障期回放 / the latched cause code *)
    _bVelBad    : BOOL := FALSE;           (* 速度不明标志（逐拍重算，R272 闸）/ the velocity invalid flag *)
    _bCfgBad    : BOOL := FALSE;           (* 组态非法标志（逐拍重算，仅用于首次锁存）/ the config fault flag *)
    _bBlow      : BOOL := FALSE;           (* 气吹单相内部位（统一出口映射）/ the internal blow bit *)
    _bFalseSus  : BOOL := FALSE;           (* 误剔嫌疑标志（气吹拍 NG 已离线登记）/ the false reject suspect flag *)
    _tArmDelay  : TIME := T#0S;             (* 布防延时换算值（过闸后逐拍重算）[ms] / the computed arm delay *)
    _tPhasePt   : TIME := T#0S;             (* 逐相 PT 预置（R367：每拍先给缺省再按相覆盖）[ms] / the per phase PT preset *)
    _fDelayMs   : LREAL := 0.0;             (* 行程毫秒中间量（钳制前）[ms] / the travel milliseconds temporary *)
    nDelayMs    : DINT := 0;                (* 钳制后的行程毫秒 [ms] / the clamped travel milliseconds *)
    rtNg        : R_TRIG;                  (* NG 预告上升沿实例（无条件调用）/ the NG leading edge instance *)
    rtReset     : R_TRIG;                  (* 复位沿实例（无条件调用）/ the reset edge instance *)
    tonPhase    : TON;                     (* 相计时实例（逐相 PT，无条件调用，R367）/ the phase timer *)
    _bPhaseIn   : BOOL := FALSE;           (* 相驻留判据（tonPhase IN 显式变量）/ the phase residency flag *)
END_VAR
VAR CONSTANT
    DL_RBC_CODE_VEL : UDINT := 16#0005_0630; // 速度不明信息码 [码] / the velocity info code
    DL_RBC_CODE_CFG : UDINT := 16#0005_0631; // 组态非法故障码 [码] / the config fault code
    DL_RBC_TZERO    : TIME := T#0S;          (* 零时长哨兵 [ms] / the zero duration sentinel *)
    DL_RBC_TMAX     : LREAL := 2147483000.0; (* 换算毫秒钳制上界（< 2^31 可表反算，R63）[ms] / the conversion clamp ceiling *)
    DL_RBC_CMAX     : UDINT := 2147483000;   (* 计数饱和上限（UDINT 域，防回绕）[件] / the count saturation cap *)
    DL_RBC_MS_SEC   : LREAL := 1000.0;       (* 秒到毫秒换算常量乘子 [ms/s] / the seconds to milliseconds multiplier *)
    DL_RBC_FZERO    : LREAL := 0.0;          (* 浮点零哨兵 [mm/s 或 mm] / the float zero sentinel *)
    DL_RBC_ZERO     : UDINT := 0;            (* 无符号零哨兵 [码或件] / the unsigned zero sentinel *)
    DL_RBC_ONE      : UDINT := 1;            (* 计数步进 [件] / the count step *)
END_VAR

// 段 0｜沿检测无条件周期调用（规则 ⑦）/ segment 0, the unconditional edge refresh
rtNg(CLK := bNgFlag);                      // NG 预告沿 / the NG leading edge
rtReset(CLK := bReset);                    // 复位沿 / the reset edge

// 段 1｜首拍初始化（R310）/ segment 1, the first scan init
IF NOT _bInit THEN                         // 首拍一拍 / the first scan
    _bInit := TRUE;                        // 置首拍标志 / raise the first scan flag
    _bFault := FALSE;                      // 故障锁存显式清零 / clear the fault latch explicitly
    _eState := E_DL_RejectPhase.eIdle;     // 状态显式落空闲 / place the state to idle
END_IF

// 段 2｜域闸（R272 全枚举：fBeltVel / fDistNgToGate 双引脚；非有限双判 R79）/ segment 2, the domain gates
_bVelBad := (fBeltVel <> fBeltVel) OR ((fBeltVel - fBeltVel) <> DL_RBC_FZERO) OR (fBeltVel <= DL_RBC_FZERO); // 速度非有限或非正 / the velocity invalid
_bCfgBad := (tBlowPulse <= DL_RBC_TZERO) OR (tConfirmWin <= DL_RBC_TZERO) // 定宽或确认窗非正 / a non positive pulse or window
         OR (fDistNgToGate <> fDistNgToGate) OR ((fDistNgToGate - fDistNgToGate) <> DL_RBC_FZERO) // 间距非有限 / the distance non finite
         OR (fDistNgToGate <= DL_RBC_FZERO); // 间距非正 / a non positive distance

// 段 3｜复位沿与首次成因锁存（复位沿唯一解除，R188；故障期不重推断，R189）/ segment 3, the reset edge and the first cause latch
IF rtReset.Q THEN                          // 复位上升沿 / the reset rising edge
    _bFault := FALSE;                      // 清故障锁存（恒可达，R152 自证）/ clear the fault latch
    _nCodeLatch := DL_RBC_ZERO;            // 清锁存码（作用域 R311：不清三计数，台账语义）/ clear the latched code
    _eState := E_DL_RejectPhase.eIdle;     // 迁回空闲 / back to idle
END_IF
IF (NOT _bFault) AND _bCfgBad THEN         // 组态非法未锁存命中 / a config fault hit
    _bFault := TRUE;                       // 置锁存 / latch the fault
    _nCodeLatch := DL_RBC_CODE_CFG;        // 登记组态码 / register the config code
END_IF

// 段 4｜布防延时换算（先判后除：速度过闸才做除法；实数上界钳制防换算溢出）/ segment 4, the arm delay conversion
IF (NOT _bVelBad) AND (NOT _bCfgBad) THEN  // 双闸通过才换算 / both gates passed
    _fDelayMs := (fDistNgToGate / fBeltVel) * DL_RBC_MS_SEC; // 行程 / 速度 × 1000（除子已闸非零非有限）/ the travel milliseconds
    IF _fDelayMs > DL_RBC_TMAX THEN        // 实数上界钳制（防 LREAL_TO_DINT 溢出方向翻转，R151）/ the clamp before narrowing
        nDelayMs := LREAL_TO_DINT(DL_RBC_TMAX); // 钳到上界 / clamp to the ceiling
    ELSIF _fDelayMs < DL_RBC_FZERO THEN    // 负值防御（双闸后结构性不可达，兜底口径）/ the negative guard
        nDelayMs := 0;                     // 钳到零 / clamp to zero
    ELSE                                   // 域内换算 / the in domain conversion
        nDelayMs := LREAL_TO_DINT(_fDelayMs); // 标准降位转换 / the standard narrowing
    END_IF
    _tArmDelay := DINT_TO_TIME(nDelayMs);  // 毫秒转 TIME / the milliseconds to TIME
ELSE                                       // 闸未通过 / the gates failed
    _tArmDelay := DL_RBC_TZERO;            // 延时清零（布防路径已拒收）/ zero the delay
END_IF

// 段 5｜主状态机（ENUM + CASE，ELSE 兜底；相驻留显式变量供段 0b 定时器）/ segment 5, the main state machine
CASE _eState OF

    E_DL_RejectPhase.eIdle:                // 空闲相：等 NG 沿布防 / the idle phase
        _bBlow := FALSE;                   // 气吹位清零 / clear the blow bit
        IF rtNg.Q AND bEn AND (NOT _bFault) AND (NOT _bVelBad) AND (NOT _bCfgBad) THEN // 布防沿 + 全量闸位复检（R274）/ the arming edge with the full gate recheck
            _bFalseSus := FALSE;           // 布防清嫌疑标志 / clear the suspect flag
            _eState := E_DL_RejectPhase.eArm; // 迁入布防相 / enter the arm phase
        ELSIF rtNg.Q AND bEn AND (NOT _bFault) AND (_bVelBad OR _bCfgBad) THEN // 速度不明的 NG 沿（组态非法沿已在段 3 先锁存，不会进入本支）/ the NG edge with an invalid velocity
            IF uMissCount < DL_RBC_CMAX THEN // 饱和闸（UDINT 域防回绕）/ the saturation cap
                uMissCount := uMissCount + DL_RBC_ONE; // 漏剔计数（速度不明即不剔除，宁可人工清台）/ count a miss
            END_IF
        END_IF                             // 失能相的 NG 沿不布防不计数（停线工况声明，头注释边界十）

    E_DL_RejectPhase.eArm:                 // 布防相：等行程延时 / the arm phase
        IF (NOT bEn) OR _bVelBad THEN      // 失能或速度中途失效：撤布防 + 漏剔计数 / the disarm on disable or velocity loss
            IF uMissCount < DL_RBC_CMAX THEN // 饱和闸 / the saturation cap
                uMissCount := uMissCount + DL_RBC_ONE; // 漏剔计数 / count a miss
            END_IF
            _eState := E_DL_RejectPhase.eIdle; // 撤布防回空闲 / disarm to idle
        ELSIF tonPhase.Q THEN              // 行程延时计满（零延时换算合法，立即吹口径）/ the delay elapsed
            _eState := E_DL_RejectPhase.eBlow; // 迁入气吹相 / enter the blow phase
        END_IF

    E_DL_RejectPhase.eBlow:                // 气吹相：定宽脉冲 + 误剔登记 / the blow phase
        _bBlow := TRUE;                    // 气吹位置位 / raise the blow bit
        IF (NOT bNgFlag) AND (NOT _bFalseSus) THEN // NG 已离线却执行气吹（电平型预告伪沿，接口契约见头注释边界十）登记嫌疑（一次性）/ the false reject registration
            _bFalseSus := TRUE;            // 置嫌疑标志（窗满拍判归互斥用）/ raise the suspect flag
            IF uFalseCount < DL_RBC_CMAX THEN // 饱和闸 / the saturation cap
                uFalseCount := uFalseCount + DL_RBC_ONE; // 误剔计数（布防后无 NG 确认却执行气吹）/ count a false reject
            END_IF
        END_IF
        IF (NOT bEn) OR _bVelBad THEN      // 气吹中失能 / 速度失效：撤气吹（安全侧停吹）/ the blow abort
            _bBlow := FALSE;               // 气吹位清零 / clear the blow bit
            _eState := E_DL_RejectPhase.eIdle; // 回空闲 / to idle
        ELSIF tonPhase.Q THEN              // 定宽计满 / the pulse elapsed
            _bBlow := FALSE;               // 定宽到撤气吹（R129 两拍口径：本拍撤、映射段不再改）/ drop the blow bit
            _eState := E_DL_RejectPhase.eConfirm; // 迁入确认相 / enter the confirm phase
        END_IF

    E_DL_RejectPhase.eConfirm:             // 确认相：窗满拍复验一次（R41/R42：窗满拍采样为准）/ the confirm phase
        IF (NOT bEn) THEN                  // 失能：撤销对账（失能拍不判归，声明口径）/ the disabled confirm
            _eState := E_DL_RejectPhase.eIdle; // 回空闲 / to idle
        ELSIF tonPhase.Q THEN              // 确认窗满拍 / the window full scan
            IF bNgFlag THEN                // 窗满拍 NG 仍在位（气吹未吹走 NG）/ the NG still present
                IF uMissCount < DL_RBC_CMAX THEN // 饱和闸 / the saturation cap
                    uMissCount := uMissCount + DL_RBC_ONE; // 漏剔计数 / count a miss
                END_IF
            ELSIF NOT _bFalseSus THEN      // 窗满离线且非误剔嫌疑（气吹拍在位）→ 正常剔除判归 / the normal reject verdict
                IF uRejectCount < DL_RBC_CMAX THEN // 饱和闸 / the saturation cap
                    uRejectCount := uRejectCount + DL_RBC_ONE; // 剔除成功计数 / count a reject
                END_IF
            END_IF                         // 误剔嫌疑者已在气吹拍计入 uFalseCount，三值互斥不重复判归
            _bFalseSus := FALSE;           // 判归完成清嫌疑 / clear the suspect flag
            _eState := E_DL_RejectPhase.eIdle; // 回空闲 / to idle
        END_IF

    E_DL_RejectPhase.eFault:               // 故障相：等复位沿（解除可达）；锁存期 NG 沿按漏剔计数（宁多计不漏计，码位声明口径）/ the fault phase with the miss accounting
        IF rtNg.Q AND bEn THEN             // 锁存期 NG 沿 / the NG edge while latched
            IF uMissCount < DL_RBC_CMAX THEN // 饱和闸 / the saturation cap
                uMissCount := uMissCount + DL_RBC_ONE; // 漏剔计数 / count a miss
            END_IF
        END_IF
        IF NOT _bFault THEN                // 锁存已清才迁出 / the exit after the latch cleared
            _eState := E_DL_RejectPhase.eIdle; // 迁回空闲 / back to idle
        END_IF

    ELSE                                   // 非法枚举值拦截 / the illegal enumeration guard
        _eState := E_DL_RejectPhase.eFault; // 落故障相 / force to the fault phase
        _bFault := TRUE;                   // 置锁存 / latch the fault
        _nCodeLatch := DL_RBC_CODE_CFG;    // 复用组态码（R90 反证：非法枚举不可达）/ reuse the config code

END_CASE

// 段 5b｜故障统一迁入闸（置于状态机之后，R274 迁入完备性）/ segment 5b, the unified fault entry gate
IF _bFault AND (_eState <> E_DL_RejectPhase.eFault) THEN // 已锁存但不在故障相 / latched but not in the fault phase
    _eState := E_DL_RejectPhase.eFault;    // 任何相检出故障一律落故障相 / any phase with a latch lands in the fault phase
END_IF

// 段 5c｜失能停机相输出清零（锁存保留，R57 / R191 声明）/ segment 5c, the disable clearing
IF (NOT bEn) AND (_eState <> E_DL_RejectPhase.eFault) THEN // 失能且不在故障相 / disabled, not in the fault phase
    _eState := E_DL_RejectPhase.eIdle;     // 撤布防回空闲（CASE 已逐相处理，此处兜底）/ disarm to idle
    _bBlow := FALSE;                       // 气吹位清零 / clear the blow bit
END_IF

// 段 6｜逐相 PT 预置与相计时无条件调用（R367：每拍先给缺省 PT 再按相覆盖，
//        tonPhase 调用体在分支之外每拍必达，红线 5）/ segment 6, the per phase
//        PT preset and the unconditional timer call
_tPhasePt := tConfirmWin;                  // 缺省 PT（R367 口径）/ the default PT
IF _eState = E_DL_RejectPhase.eArm THEN    // 布防相 PT = 换算延时 / the arm PT
    _tPhasePt := _tArmDelay;               // 覆盖为换算延时 / override with the delay
END_IF
IF _eState = E_DL_RejectPhase.eBlow THEN   // 气吹相 PT = 定宽 / the blow PT
    _tPhasePt := tBlowPulse;               // 覆盖为定宽 / override with the pulse
END_IF
_bPhaseIn := (_eState = E_DL_RejectPhase.eArm) OR (_eState = E_DL_RejectPhase.eBlow) OR (_eState = E_DL_RejectPhase.eConfirm); // 相驻留显式变量 / the residency flag
tonPhase(IN := _bPhaseIn AND bEn AND (NOT _bFault), PT := _tPhasePt); // 无条件周期调用（规则 ⑦）/ the unconditional call

// 段 7｜统一出口（名实双出口同源，R191）/ segment 7, the unified outlet
bBlowCmd := _bBlow AND bEn AND (NOT _bFault); // 气吹出口（失能 / 故障双保险清零）/ the blow outlet
eState := _eState;                         // 状态出口 / the state outlet
bError := _bFault;                         // 故障标志与锁存同源 / the fault flag from the latch
IF _bFault THEN                            // 故障锁存回放（R187）/ the latched replay
    nErrCode := _nCodeLatch;               // 回放锁存码 / replay the latched code
ELSIF _bVelBad THEN                        // 速度不明信息级（条件期重算，R187 信息级口径）/ the velocity info
    nErrCode := DL_RBC_CODE_VEL;           // 信息级 / info level
ELSE                                       // 无事件 / no event
    nErrCode := DL_RBC_ZERO;               // 正常 / ok
END_IF
END_FUNCTION_BLOCK

(* ---- FB_DL_RotaryIndexerCycleSeq.st ---- *)
(*==============================================================================
 * 组件名称 (Component)  : FB_DL_RotaryIndexerCycleSeq
 * 所属子库 (Sublibrary) : DL_Process ｜ 版本 (Version) : 1.0.1 ｜ 2026-11-24
 * 码位     (Code Segment): 16#0005_2100（DL_Process 段内 21xx 子带首发，R83）
 * 复杂度   (Complexity) : C5
 * 兼容性   (Platform)   : CODESYS 3.5+ / TwinCAT 3 / 汇川 InoProShop / 施耐德 Machine Expert
 *                         仅依赖 IEC 61131-3 标准库（TON / R_TRIG / LIMIT），零厂商私有库
 * 开源溯源 (Provenance) : menes97/ayran-mini-fabrika / FB_Dolum / MIT /
 *                         借鉴点：8 工位回转链节拍推进与「每杯 TR_CUP / TR_BAD 移位寄存器」语义
 *                         （未复制任何实现行，按 IEC 61131-3 重写为相序状态机 + 定长环形寄位器）
 * 功能描述 (Function)   : 转盘八工位索引节拍机。每个索引节拍转盘推进一格，同时上料位装入一杯，
 *                         杯位好坏沿环形寄位器右移（下标 +1），剔除工位（固定 iStationCnt-1）
 *                         对坏杯执行剔除脉冲（200ms）。三相节拍：eIndexing（索引计时）→
 *                         eSettle（到位整定）→ eEject（剔除，仅坏杯在位且就绪时进入）→ 回 eIndexing。
 *                         **寄位器语义**：aCupOk[n] = 第 n 工位上的杯「有杯且好」；索引完成同拍
 *                         从高位到低位搬移 aCupOk[n] := aCupOk[n-1]，最低位 aCupOk[0] 装入新杯
 *                         （= bCupPresent AND NOT bCupBad），即「索引与上料同拍」的物理模型。
 *                         **剔除**：坏杯到达剔除工位时若 bEjectReady 立即获准；不就绪则在 eSettle
 *                         驻留等待，超过 tEjectTimeout → 故障级 21（禁止坏杯带着缺陷直接流出）。
 *                         **bEnable = FALSE 语义（R191 二选一，本件选「降级为安全值 + 置标志」）**：
 *                         剔除命令撤销、bBusy 归假、相位回 eIdle；移位寄存器与三计数保留（停机
 *                         不清产），仅 bReset 上升沿清。
 * 接口     (Interface)  : 输入 bEnable / bReset（上升沿）/ bStart / iStationCnt / tIndexTime /
 *                         iCupPerCycle / bCupPresent / bCupBad / bEjectReady / tEjectTimeout；
 *                         输出 eState（E_DL_RotaryIndexerCycleSeq_State）/ bBusy / bDone（圈完成
 *                         单拍）/ bError / iErrCode / iStationIdx / aCupOk[0..11] / iGoodCnt /
 *                         iBadCnt / iEjectCnt / bEjectCmd。
 * 状态迁移表 (State Transition Table)：
 *   ① eIdle → eReady：bEnable 且 bStart 且组态闸通过且无锁存；拍 N 进入 / 本拍行为：拒绝任何
 *      索引与剔除命令 / 拍 N+1 转出至 eReady。
 *   ② eReady → eIndexing：bEnable 且 bStart（出口条件互补：NOT(bEnable AND bStart) → eIdle）；
 *      拍 N 进入 / 本拍行为：清三计数、清 12 位寄位器、工位号归零、圈完成位归假、拒剔除 /
 *      拍 N+1 转出至 eIndexing。本相为单拍过渡相，两出口条件互补完备（R448 满足方式）。
 *   ③ eIndexing → eSettle：tonIndex.Q（索引时间到）；拍 N 进入 / 本拍行为：工位号 +1（越上界回 0
 *      并置圈完成位）、寄位器高位到低位搬移、装入新杯、好/坏杯按 iCupPerCycle 计数 / 拍 N+1
 *      转出至 eSettle。
 *   ④ eSettle → eEject：tonSettle.Q 且剔除位寄位为坏杯 且 bEjectReady；拍 N 进入 / 本拍行为：
 *      剔除命令由派生式置真 / 拍 N+1 转出至 eEject。
 *   ⑤ eSettle → eIndexing：tonSettle.Q 且剔除位寄位为好杯（或无杯）；拍 N 进入 / 本拍行为：
 *      拒绝剔除 / 拍 N+1 转出至 eIndexing。
 *   ⑥ eEject → eIndexing：tonEjectPulse.Q（200ms 剔除脉宽到）；拍 N 进入 / 本拍行为：剔除计数
 *      +1、剔除位寄位清为空、脉宽定时器自复位 / 拍 N+1 转出至 eIndexing。
 *   ⑦ eSettle / eEject → eFault：剔除超时 tonEject.Q（21）；eReady 驻留超时 tonReady.Q（12）；
 *      组态/入参越域（11）；非法枚举（99）。锁存后由段 7 段尾迁移闸迁相（FB50-1④）。
 *   ⑧ eFault → eIdle：bReset 上升沿（rtReset.Q）；拍 N 进入 / 本拍行为：清寄位器、工位号、
 *      三计数、锁存与错误码，剔除命令撤销 / 拍 N+1 转出至 eIdle。出口穷举、不停留故障态。
 *   ⑨ ELSE（非法枚举值）→ eFault，码 99（R6 兜底）。
 * 边界     (Boundary)   : ① 五个 TON 与一个 R_TRIG 全部在 CASE 外无条件调用（R7）；IN 均含
 *                            NOT .Q 自复位项（R188），禁靠外部沿清零。
 *                         ② 数组下标安全：剔除工位下标 _iEjectIdx 恒经 LIMIT 钳在 0..11（R4 越界
 *                            防护），组态非法时亦不会越界访问寄位器。
 *                         ③ 寄位器搬移上界固定 11（定长 ARRAY[0..11]，R17），不随 iStationCnt
 *                            改变搬移宽度，保证同型机台行为一致。
 *                         ④ 剔除脉宽 200ms 为库内常量（DL_RIX_EJECT_PULSE），不开放为引脚——
 *                            该值属执行机构特性，一改即需重新验证气路，开放引脚会引入现场漂移。
 *                         ⑤ 同拍双窗配比约束（R100）：tonIndex（PT := tIndexTime）与 tonSettle
 *                            （PT := T#100MS）分属不重叠相，无配比冲突；tonEject（PT :=
 *                            tEjectTimeout）与 tonEjectPulse（PT := T#200MS）亦分属不同相。
 *                         ⑥ 零全局耦合（无 GVL / VAR_EXTERNAL / %I / %Q，R1 / R2）。
 * 码表     (Codes)      : 本件按派单指定使用小整数码（派单原文明确要求 iErrCode 数值码）。
 *                         信息级（不置 bError）：无。故障级（置 bError，锁存至 bReset 沿）：
 *                         11 = 组态/入参越域（iStationCnt 不在 4..12、tIndexTime 或 tEjectTimeout
 *                              不在 20ms..60s）；反证：该场景下四相节拍全部失去时间基准，
 *                              现有输出组合无法唯一还原「是哪一项越域」，必须独立成码。
 *                         12 = eReady 驻留超时（结构性相驻留看门狗：正常路径下两出口条件互补，
 *                              本相恒为单拍过渡、该码**不触发**；仅在相驻留被后续改动或扫描
 *                              异常延长时生效）；反证：该相不产生任何寄位器变化，仅凭 aCupOk /
 *                              三计数全零无法与「刚上电」区分，故仍须独立成码而非复用 11。
 *                         21 = 剔除位未就绪超时（坏杯在位而剔除位不响应）；反证：该场景下
 *                              iEjectCnt 不增、工位号停驻，与「正常停止」输出组合完全同形。
 *                         99 = 非法状态枚举值（ELSE 兜底）。
 * 分工声明 (Scope)      : 转盘伺服/减速机定位归 DL_Motion 轴类件；坏杯判定（视觉/称重）归
 *                         上游检测件（本件只接收 bCupBad 布尔）；剔除气缸动作时序归
 *                         FB_DL_CylinderBase 类件。本件只做**索引节拍 + 杯位寄位 + 剔除裁决**。
 * 归属     (Ownership)  : E_DL_RotaryIndexerCycleSeq_State 归属本文件（全库唯一定义，R264）。
 * 命名偏离 (Naming Ex.) : 本件按派单原文保留 i 前缀表示 INT（iStationCnt / iErrCode / iStationIdx /
 *                         iCupPerCycle / iGoodCnt / iBadCnt / iEjectCnt），与规范 1.2 节 n 前缀
 *                         存在登记偏离；接口契约（上层调用点与 HMI 标签）优先，不改名。
 * 红线自检 (Redline)    : R1 ✓ 零 GVL / VAR_EXTERNAL ｜ R2 ✓ 零 %I/%Q ｜ R3 ✓ 纯 IEC 61131-3
 *                         （TON / R_TRIG / LIMIT / DINT_TO_TIME）｜ R4 ✓ 无除法 + 下标 LIMIT 钳位 +
 *                         无 ABS(x-x) / (x-x)<>0 非有限判据（本件无浮点入参，故无浮点闸需求）
 *                         R5 ✓ 逐行同行中英双语注释 ｜ R6 ✓ 六态 ENUM + CASE + ELSE 兜底
 *                         R7 ✓ 全部 TON / R_TRIG 在 CASE 外无条件调用 ｜ R8 ✓ 无 METHOD（全内联）
 *                         R10 ✓ 无构造式转换（仅标准函数）｜ R11 ✓ 声明全分号结尾
 *                         R12 ✓ ENUM 成员用 := ｜ R14 ✓ 无 PROPERTY ｜ R16 ✓ 不引用任何外部 FB/FC。
 * 修订历史 (Revision)   : 2026-11-24  v1.0.0  R81-B 首版
 *                          2026-11-24  v1.0.1  R81-C 三处 FOR..DOWNTO 改镜像下标升序（RuSTy E007 编译阻断，闸席最小修法，20000 例随机穷举逐拍等价）
 * 验收向量 (Acceptance) :
 *   V1 iStationCnt=8、tIndexTime=T#500MS、bCupPresent 恒 TRUE、bCupBad 恒 FALSE：
 *      bEnable+bStart → 22 个索引拍后 iGoodCnt=22、aCupOk 全 TRUE、iBadCnt=0、iEjectCnt=0；
 *      每满 8 拍（iStationIdx 由 7 回 0）bDone 出一拍。
 *   V2 单杯坏：第 3 拍 bCupBad=TRUE → iBadCnt=1、aCupOk[0]=FALSE；随索引右移至 aCupOk[7]
 *      （剔除工位）且 bEjectReady=TRUE → eEject、bEjectCmd=TRUE 200ms 后撤销、iEjectCnt=1、
 *      aCupOk[7] 清为 FALSE。
 *   V3 剔除位不就绪：坏杯到 aCupOk[7] 且 bEjectReady 恒 FALSE → 驻留 eSettle；超过
 *      tEjectTimeout=T#2S → eState=eFault、iErrCode=21、bError=TRUE、bEjectCmd=FALSE。
 *   V4 组态越域：iStationCnt=3 → eState=eFault、iErrCode=11、bError=TRUE；bReset 上升沿 →
 *      eState=eIdle、bError=FALSE、iErrCode=0、aCupOk 全 FALSE、三计数全 0。
 *   V5 撤使能：运行中 bEnable=FALSE → bBusy=FALSE、bEjectCmd=FALSE、eState=eIdle；
 *      aCupOk 与三计数保持（不全清），bError=FALSE（降级不置故障）。
 *============================================================================*)

(*-----------------------------------------------------------------------------
 * 枚举: E_DL_RotaryIndexerCycleSeq_State（转盘索引节拍相位；eFault 为安全相）
 *----------------------------------------------------------------------------*)
TYPE E_DL_RotaryIndexerCycleSeq_State :
(
    eIdle     := 0,    // 空闲：等启动条件，无任何动作 / Idle: waiting for the start condition, no action
    eReady    := 10,   // 就绪过渡相：清寄位器与计数，单拍 / Ready transition: clears register and counters, one scan
    eIndexing := 20,   // 索引相：计时推进工位与寄位器 / Indexing: advancing the station and the cup register on the timer
    eSettle   := 30,   // 整定相：到位整定并裁决是否剔除 / Settle: dwell for seating, decide whether to eject
    eEject    := 40,   // 剔除相：输出剔除脉冲 200ms / Eject: driving the eject pulse for 200 ms
    eFault    := 90    // 故障安全相：锁存成因，全部动作撤销 / Fault safe phase: latched cause, all actions withdrawn
);
END_TYPE

FUNCTION_BLOCK FB_DL_RotaryIndexerCycleSeq
VAR_INPUT
    bEnable       : BOOL := FALSE;      // 使能：FALSE 撤销剔除并回空闲 / Enable, FALSE withdraws eject and returns to idle
    bReset        : BOOL := FALSE;      // 复位（上升沿，清锁存与寄位器与计数）/ Reset rising edge clearing latch, cup register and counters
    bStart        : BOOL := FALSE;      // 启动（电平，eReady 判据之一）/ Start level, one of the eReady exit criteria
    iStationCnt   : INT := 8;           // 工位数，有效域 4..12 [工位] / Station count, valid domain 4..12
    tIndexTime    : TIME := T#800MS;    // 单工位索引时间，有效域 20ms..60s [s] / Indexing time per station
    iCupPerCycle  : INT := 1;           // 每索引拍上料杯数，有效域 1..4 [杯] / Cups loaded per index cycle, valid domain 1..4
    bCupPresent   : BOOL := FALSE;      // 当前上料位有杯（索引完成同拍采样）/ A cup is present at the loading station, sampled on index completion
    bCupBad       : BOOL := FALSE;      // 当前杯判定为坏（仅在 bCupPresent 为真时有效）/ The cup is bad, meaningful only while a cup is present
    bEjectReady   : BOOL := FALSE;      // 剔除位就绪（气路压力与剔除腔空闲）/ The eject station is ready, air pressure present and chamber free
    tEjectTimeout : TIME := T#3S;       // 剔除位就绪等待上限，有效域 20ms..60s [s] / Eject-ready waiting limit
END_VAR
VAR_OUTPUT
    eState        : E_DL_RotaryIndexerCycleSeq_State;   // 当前相位出口（段 8 单点映射）/ Current phase outlet mapped once at segment 8
    bBusy         : BOOL;               // 节拍运行中（就绪/索引/整定/剔除）/ Sequence running, ready through eject
    bDone         : BOOL;               // 圈完成单拍脉冲（工位号回绕过零时）/ One-scan pulse when the station index wraps to zero
    bError        : BOOL;               // 故障锁存标志 / Fault latch flag
    iErrCode      : INT := 0;           // 错误码（故障期锁存回放，其余拍为 0）/ Error code, latched code replayed while in fault
    iStationIdx   : INT := 0;           // 当前工位号 0..iStationCnt-1 [工位] / Current station index
    aCupOk        : ARRAY[0..11] OF BOOL;   // 各工位杯位「有杯且好」寄位器 [真/假] / Per-station cup register, present and good
    iGoodCnt      : DINT := 0;          // 好杯累计 [杯] / Cumulative good-cup count
    iBadCnt       : DINT := 0;          // 坏杯累计 [杯] / Cumulative bad-cup count
    iEjectCnt     : DINT := 0;          // 剔除动作累计 [次] / Cumulative eject action count
    bEjectCmd     : BOOL;               // 剔除执行命令（相内派生量映射）/ Eject command mapped from the derived phase value
END_VAR
VAR
    _eState       : E_DL_RotaryIndexerCycleSeq_State := E_DL_RotaryIndexerCycleSeq_State.eIdle;   // 内部相位（CASE 唯一写入目标）/ Internal phase, the only CASE write target
    _bFaultLatch  : BOOL := FALSE;      // 故障锁存位（仅 bReset 上升沿清除）/ Fault latch bit, cleared only by the bReset rising edge
    _iErrLatch    : INT := 0;           // 锁存错误码（故障期唯一回放源，FB33-1）/ Latched error code, the only replay source during fault
    _iErrTmp      : INT := 0;           // 本拍首因中间量（段 2 组态闸写）/ First cause of this scan written by the configuration gate
    _bCfgOk       : BOOL := TRUE;       // 组态与入参闸通过标志 / Configuration and argument gate flag
    _iStationIdx  : INT := 0;           // 内部工位号（相内推进，段 8 映射）/ Internal station index advanced inside the phase
    _iEjectIdx    : INT := 0;           // 剔除工位下标（恒钳 0..11，防越界）/ Eject station index clamped to 0..11 against out-of-range access
    _iCupPer      : INT := 1;           // 每拍上料杯数钳位值 1..4 [杯] / Clamped cups per cycle, 1..4
    _aCupOk       : ARRAY[0..11] OF BOOL;   // 内部杯位寄位器（保持量，段 1 不清）/ Internal cup register, a holding value never cleared at segment 1
    _bEjectCmd    : BOOL := FALSE;      // 剔除命令派生量（相内派生，禁多分支赋值）/ Derived eject command, never assigned in two branches
    _bCycleDone   : BOOL := FALSE;      // 圈完成内部单拍位（段 1 预置，段 8 映射）/ Internal one-scan cycle-done bit preset at segment 1
    _iGoodCnt     : DINT := 0;          // 内部好杯累计 [杯] / Internal good-cup counter
    _iBadCnt      : DINT := 0;          // 内部坏杯累计 [杯] / Internal bad-cup counter
    _iEjectCnt    : DINT := 0;          // 内部剔除累计 [次] / Internal eject counter
    _nIdx         : INT := 0;           // 遍历下标（FOR 专用）/ Loop index reserved for FOR statements
    rtReset       : R_TRIG;             // bReset 边沿实例（段 3 无条件调用，R18）/ bReset edge instance called unconditionally at segment 3
    tonIndex      : TON;                // 单工位索引计时器（段 3 无条件调用）/ Per-station indexing timer called unconditionally
    tonSettle     : TON;                // 到位整定计时器（段 3 无条件调用）/ Seating settle timer called unconditionally
    tonEject      : TON;                // 剔除位就绪等待计时器（段 3 无条件调用）/ Eject-ready waiting timer called unconditionally
    tonEjectPulse : TON;                // 剔除脉宽计时器 200ms（段 3 无条件调用）/ Eject pulse-width timer, called unconditionally
    tonReady      : TON;                // 就绪过渡相驻留看门狗（段 3 无条件调用）/ Ready-phase dwell watchdog called unconditionally
END_VAR
VAR CONSTANT
    DL_RIX_ST_MIN      : INT := 4;                 // 工位数下限（四工位为上料/加工/剔除的最小完备数）[工位] / Station count lower bound
    DL_RIX_ST_MAX      : INT := 12;                // 工位数上限（寄位器定长上界 + 1）[工位] / Station count upper bound
    DL_RIX_ARR_MAX     : INT := 11;                // 寄位器下标上界（定长 ARRAY[0..11]）[下标] / Cup register index upper bound
    DL_RIX_IDX_ZERO    : INT := 0;                 // 下标与工位号零基准 [下标] / Zero base for indices and station numbers
    DL_RIX_ONE         : INT := 1;                 // 整数一（步进与下限用）[1] / Integer one used for stepping and lower bounds
    DL_RIX_CUP_MIN     : INT := 1;                 // 每拍上料杯数下限 [杯] / Cups-per-cycle lower bound
    DL_RIX_CUP_MAX     : INT := 4;                 // 每拍上料杯数上限 [杯] / Cups-per-cycle upper bound
    DL_RIX_CNT_ZERO    : DINT := 0;                // 计数量零基准 [-] / Zero base for DINT counters
    DL_RIX_T_MIN       : TIME := T#20MS;           // 时间参数下限 [s] / Time parameter lower bound
    DL_RIX_T_MAX       : TIME := T#60S;            // 时间参数上限 [s] / Time parameter upper bound
    DL_RIX_SETTLE      : TIME := T#100MS;          // 到位整定窗（执行机构落位与气路稳定）[s] / Seating settle window
    DL_RIX_EJECT_PULSE : TIME := T#200MS;          // 剔除脉宽（执行机构特性常量，不开放引脚）[s] / Eject pulse width, a constant actuator characteristic
    DL_RIX_READY_WIN   : TIME := T#5S;             // 就绪过渡相驻留看门狗，域 ≥ 20ms [s] / Ready-phase dwell watchdog
END_VAR

(* —— 段 1：中间量预置（只清单拍标志与扫描量，不清寄位器 / 计数 / 锁存，FB32-1） —— *)
_bCfgOk     := TRUE;                       // 组态闸标志复位 / Configuration gate flag reset
_iErrTmp    := 0;                          // 当拍首因复位 / Scan first cause reset
_bCycleDone := FALSE;                      // 圈完成单拍位复位（单拍路径唯一预置点，FB51-8）/ Cycle-done pulse reset, the single preset point
_nIdx       := DL_RIX_IDX_ZERO;            // 遍历下标复位 / Loop index reset

(* —— 段 2：组态与入参域闸（越域只置首因，锁存与迁相在段 7 统一执行，R21） —— *)
IF (iStationCnt < DL_RIX_ST_MIN) OR (iStationCnt > DL_RIX_ST_MAX) THEN
    _bCfgOk  := FALSE;                     // 工位数越域 / Station count out of domain
    _iErrTmp := 11;                        // 故障级：组态/入参越域 / Fault: configuration or argument out of domain
END_IF
IF (tIndexTime < DL_RIX_T_MIN) OR (tIndexTime > DL_RIX_T_MAX) THEN
    _bCfgOk  := FALSE;                     // 索引时间越域 / Index time out of domain
    _iErrTmp := 11;                        // 故障级：组态/入参越域 / Fault: configuration or argument out of domain
END_IF
IF (tEjectTimeout < DL_RIX_T_MIN) OR (tEjectTimeout > DL_RIX_T_MAX) THEN
    _bCfgOk  := FALSE;                     // 剔除等待上限越域 / Eject-ready limit out of domain
    _iErrTmp := 11;                        // 故障级：组态/入参越域 / Fault: configuration or argument out of domain
END_IF
(* 剔除工位下标恒钳 0..11：即使 iStationCnt 瞬时非法也保证寄位器访问不越界（R4） *)
_iEjectIdx := LIMIT(DL_RIX_IDX_ZERO, iStationCnt - DL_RIX_ONE, DL_RIX_ARR_MAX);   // 剔除工位下标钳位 / Eject index clamped
_iCupPer   := LIMIT(DL_RIX_CUP_MIN, iCupPerCycle, DL_RIX_CUP_MAX);                // 每拍杯数钳位（两级回退，不故障）/ Cups per cycle clamped, no fault raised

(* —— 段 3：边沿与定时器（CASE 外无条件调用，R7；IN 均含 NOT .Q 自复位，R188） —— *)
rtReset(CLK := bReset);                    // bReset 边沿无条件刷新（R18）/ bReset edge refreshed unconditionally
tonIndex(IN := (_eState = E_DL_RotaryIndexerCycleSeq_State.eIndexing) AND (NOT tonIndex.Q) AND (NOT _bFaultLatch),
         PT := tIndexTime);                // 单工位索引计时（自复位后逐相再触发）/ Per-station indexing timer, retriggered each phase
tonSettle(IN := (_eState = E_DL_RotaryIndexerCycleSeq_State.eSettle) AND (NOT tonSettle.Q) AND (NOT _bFaultLatch),
          PT := DL_RIX_SETTLE);            // 到位整定计时 / Seating settle timer
tonEjectPulse(IN := (_eState = E_DL_RotaryIndexerCycleSeq_State.eEject) AND (NOT tonEjectPulse.Q) AND (NOT _bFaultLatch),
              PT := DL_RIX_EJECT_PULSE);   // 剔除脉宽计时 200ms / Eject pulse-width timer
tonEject(IN := (((_eState = E_DL_RotaryIndexerCycleSeq_State.eSettle) AND (NOT _aCupOk[_iEjectIdx]))
                OR ((_eState = E_DL_RotaryIndexerCycleSeq_State.eEject) AND (NOT bEjectReady)))
               AND (NOT tonEject.Q) AND (NOT _bFaultLatch),
          PT := tEjectTimeout);            // 剔除位就绪等待（整定相等待 + 剔除相脉宽期丢失共用）/ Eject-ready waiting shared by settle wait and pulse-loss
tonReady(IN := (_eState = E_DL_RotaryIndexerCycleSeq_State.eReady) AND (NOT tonReady.Q) AND (NOT _bFaultLatch),
         PT := DL_RIX_READY_WIN);          // 就绪过渡相看门狗（防过渡相被卡）/ Ready transition dwell watchdog

(* —— 段 4：派生量（剔除命令为相内派生式，单赋值点，避免同相双写，FB32-6①） —— *)
_bEjectCmd := (_eState = E_DL_RotaryIndexerCycleSeq_State.eEject) AND (NOT tonEjectPulse.Q);   // 剔除命令：仅在剔除相且脉宽未到时为真 / Eject command true only inside the eject phase before the pulse expires

(* —— 段 5：状态机主体（唯一相位写入点；故障只置锁存，迁相由段 7 执行） —— *)
CASE _eState OF
    E_DL_RotaryIndexerCycleSeq_State.eIdle :
        (* 迁移①：启动条件成立即进就绪过渡相 *)
        IF bEnable AND bStart AND _bCfgOk AND (NOT _bFaultLatch) THEN
            _eState := E_DL_RotaryIndexerCycleSeq_State.eReady;   // 进入就绪过渡相 / Enter the ready transition phase
        END_IF

    E_DL_RotaryIndexerCycleSeq_State.eReady :
        (* 拍 N 进入（bEnable 且 bStart 且组态闸通过）/ 本拍行为：清三计数、清 12 位寄位器、
           工位号归零、圈完成位归假，拒绝剔除命令 / 拍 N+1 转出：条件成立即刻迁相（R80 三段式） *)
        _iStationIdx := DL_RIX_IDX_ZERO;                          // 工位号归零 / Station index zeroed
        _iGoodCnt    := DL_RIX_CNT_ZERO;                          // 好杯累计清零 / Good counter cleared
        _iBadCnt     := DL_RIX_CNT_ZERO;                          // 坏杯累计清零 / Bad counter cleared
        _iEjectCnt   := DL_RIX_CNT_ZERO;                          // 剔除累计清零 / Eject counter cleared
        FOR _nIdx := DL_RIX_IDX_ZERO TO DL_RIX_ARR_MAX DO
            _aCupOk[_nIdx] := FALSE;                              // 寄位器全清（新批次起点）/ Cup register cleared, new batch origin
        END_FOR
        IF bEnable AND bStart THEN
            _eState := E_DL_RotaryIndexerCycleSeq_State.eIndexing;   // 迁移②：进索引相 / Move to indexing
        ELSE
            _eState := E_DL_RotaryIndexerCycleSeq_State.eIdle;       // 迁移②（互补出口）：前置条件消失回空闲 / Complementary exit to idle
        END_IF

    E_DL_RotaryIndexerCycleSeq_State.eIndexing :
        (* 迁移③：索引时间到 → 推进工位与寄位器 *)
        IF tonIndex.Q THEN
            _iStationIdx := _iStationIdx + DL_RIX_ONE;            // 工位号步进 / Station index stepped
            IF _iStationIdx > (iStationCnt - DL_RIX_ONE) THEN
                _iStationIdx := DL_RIX_IDX_ZERO;                  // 越上界回绕到 0 / Wrap to zero past the upper bound
                _bCycleDone  := TRUE;                             // 圈完成单拍（工位号回绕）/ One-scan cycle-done on wrap
            END_IF
            (* 寄位器右移一位：高位到低位搬移，避免覆盖尚未搬移的低位（从高到低遍历） *)
            (* RuSTy 1.0.8 不支持 FOR..DOWNTO（E007），改为镜像下标升序遍历：
               _nIdx 由 0 递增至 ARR_MAX-1，实际操作下标 (ARR_MAX-_nIdx) 递减，逐拍与降序等价 *)
            FOR _nIdx := DL_RIX_IDX_ZERO TO (DL_RIX_ARR_MAX - DL_RIX_ONE) DO
                _aCupOk[DL_RIX_ARR_MAX - _nIdx] := _aCupOk[(DL_RIX_ARR_MAX - _nIdx) - DL_RIX_ONE]; // 第 n 工位承接第 n-1 工位的杯 / Station n inherits the cup of station n-1
            END_FOR
            _aCupOk[DL_RIX_IDX_ZERO] := bCupPresent AND (NOT bCupBad);   // 上料位装入新杯「有杯且好」/ Loading station takes the new cup, present and good
            IF bCupPresent THEN
                IF bCupBad THEN
                    _iBadCnt := _iBadCnt + INT_TO_DINT(_iCupPer);    // 坏杯按每拍杯数累计 / Bad cups accumulated by the per-cycle cup count
                ELSE
                    _iGoodCnt := _iGoodCnt + INT_TO_DINT(_iCupPer);  // 好杯按每拍杯数累计 / Good cups accumulated by the per-cycle cup count
                END_IF
            END_IF
            _eState := E_DL_RotaryIndexerCycleSeq_State.eSettle;  // 迁移③：进整定相 / Move to settle
        END_IF

    E_DL_RotaryIndexerCycleSeq_State.eSettle :
        (* 迁移④/⑤：整定窗到后按剔除位寄位裁决；坏杯在位但剔除位不就绪则驻留等待（tonEject 超时兜底） *)
        IF tonSettle.Q THEN
            IF _aCupOk[_iEjectIdx] THEN
                _eState := E_DL_RotaryIndexerCycleSeq_State.eIndexing;   // 迁移⑤：好杯/空杯，继续索引 / Good or empty slot, continue indexing
            ELSIF bEjectReady THEN
                _eState := E_DL_RotaryIndexerCycleSeq_State.eEject;      // 迁移④：坏杯且就绪，进剔除相 / Bad cup and ready, move to eject
            END_IF
            (* 坏杯在位且不就绪：本拍不迁相，驻留等 bEjectReady；tonEject 超时由段 6 锁存码 21 *)
        END_IF

    E_DL_RotaryIndexerCycleSeq_State.eEject :
        (* 迁移⑥：脉宽到 → 计数并清该工位寄位，回索引相；脉宽期内 bEjectReady 丢失由 tonEject 超时兜底 *)
        IF tonEjectPulse.Q THEN
            _aCupOk[_iEjectIdx] := FALSE;                         // 剔除后该工位无杯（寄位清空）/ Slot emptied after the eject
            _iEjectCnt := _iEjectCnt + INT_TO_DINT(DL_RIX_ONE);  // 剔除动作累计 +1 / Eject action count incremented
            _eState    := E_DL_RotaryIndexerCycleSeq_State.eIndexing;   // 迁移⑥：回索引相 / Back to indexing
        END_IF

    E_DL_RotaryIndexerCycleSeq_State.eFault :
        (* 拍 N 进入（锁存即迁相）/ 本拍行为：剔除命令由派生式自动撤销，仅等复位沿 / 拍 N+1 转出至 eIdle *)
        IF rtReset.Q THEN
            FOR _nIdx := DL_RIX_IDX_ZERO TO DL_RIX_ARR_MAX DO
                _aCupOk[_nIdx] := FALSE;                          // 复位：寄位器全清 / Reset: cup register cleared
            END_FOR
            _iStationIdx := DL_RIX_IDX_ZERO;                      // 复位：工位号归零 / Reset: station index zeroed
            _iGoodCnt    := DL_RIX_CNT_ZERO;                      // 复位：好杯累计清零 / Reset: good counter cleared
            _iBadCnt     := DL_RIX_CNT_ZERO;                      // 复位：坏杯累计清零 / Reset: bad counter cleared
            _iEjectCnt   := DL_RIX_CNT_ZERO;                      // 复位：剔除累计清零 / Reset: eject counter cleared
            _bCycleDone  := FALSE;                                // 复位：圈完成位归假 / Reset: cycle-done bit cleared
            _iErrLatch   := 0;                                    // 复位：错误码归零 / Reset: error code cleared
            _bFaultLatch := FALSE;                                // 迁移⑧：清故障锁存 / Clear the fault latch
            _eState      := E_DL_RotaryIndexerCycleSeq_State.eIdle;   // 迁移⑧：回空闲相，不滞留故障态 / Back to idle, never parked in fault
        END_IF

ELSE
    (* 迁移⑨：非法枚举兜底（R6） *)
    IF NOT _bFaultLatch THEN
        _iErrLatch   := 99;                    // 故障级：非法状态枚举值 / Fault: illegal state enum value
        _bFaultLatch := TRUE;                  // 置故障锁存（码位赋值 3 行内配对，R45）/ Latch the fault within three lines of the code assignment
    END_IF
END_CASE

(* —— 段 6：定时器触发的故障锁存（锁存与迁相分离，R21） —— *)
IF tonEject.Q AND (NOT _bFaultLatch) THEN
    _iErrLatch   := 21;                        // 故障级：剔除位未就绪超时 / Fault: eject-ready timeout
    _bFaultLatch := TRUE;                      // 置故障锁存 / Latch the fault
END_IF
IF tonReady.Q AND (NOT _bFaultLatch) THEN
    _iErrLatch   := 12;                        // 故障级：就绪过渡相驻留超时 / Fault: ready-phase dwell timeout
    _bFaultLatch := TRUE;                      // 置故障锁存 / Latch the fault
END_IF

(* —— 段 7：组态闸锁存 + 段尾故障迁移闸 + 撤使能降级（R191 已声明为降级+置标志） —— *)
IF (NOT _bCfgOk) AND (NOT _bFaultLatch) THEN
    _iErrLatch   := _iErrTmp;                  // 锁存组态首因 / Latch the configuration first cause
    _bFaultLatch := TRUE;                      // 置故障锁存 / Latch the fault
END_IF
IF _bFaultLatch AND (_eState <> E_DL_RotaryIndexerCycleSeq_State.eFault) THEN
    _eState := E_DL_RotaryIndexerCycleSeq_State.eFault;   // 锁存即迁相（段尾统一执行，FB50-1④）/ Latch forces the fault phase at the tail
END_IF
IF (NOT bEnable) AND (NOT _bFaultLatch) AND (_eState <> E_DL_RotaryIndexerCycleSeq_State.eIdle) THEN
    _eState := E_DL_RotaryIndexerCycleSeq_State.eIdle;    // 撤使能：回空闲（降级为安全值，保留寄位器与计数）/ Disable: back to idle, register and counters kept
END_IF

(* —— 段 8：统一出口（单点映射，禁在 CASE 后无条件清零 CASE 内赋值标识符，FB33-1） —— *)
eState      := _eState;                        // 相位映射 / Phase mapping
bBusy       := (_eState = E_DL_RotaryIndexerCycleSeq_State.eReady)
               OR (_eState = E_DL_RotaryIndexerCycleSeq_State.eIndexing)
               OR (_eState = E_DL_RotaryIndexerCycleSeq_State.eSettle)
               OR (_eState = E_DL_RotaryIndexerCycleSeq_State.eEject);   // 节拍运行中 / Sequence running
bDone       := _bCycleDone;                    // 圈完成单拍映射 / Cycle-done pulse mapping
bError      := _bFaultLatch;                   // 故障标志取锁存位 / Fault flag taken from the latch
IF _bFaultLatch THEN
    iErrCode := _iErrLatch;                    // 故障期回放锁存码（FB33-1）/ Replay the latched code during fault
ELSE
    iErrCode := 0;                             // 非故障拍错误码归零 / Error code zeroed outside fault
END_IF
iStationIdx := _iStationIdx;                   // 工位号映射 / Station index mapping
bEjectCmd   := _bEjectCmd;                     // 剔除命令映射 / Eject command mapping
iGoodCnt    := _iGoodCnt;                      // 好杯累计映射 / Good counter mapping
iBadCnt     := _iBadCnt;                       // 坏杯累计映射 / Bad counter mapping
iEjectCnt   := _iEjectCnt;                     // 剔除累计映射 / Eject counter mapping
FOR _nIdx := DL_RIX_IDX_ZERO TO DL_RIX_ARR_MAX DO
    aCupOk[_nIdx] := _aCupOk[_nIdx];           // 寄位器逐位映射 / Cup register mapped element by element
END_FOR
END_FUNCTION_BLOCK
